Fanuc KAREL source: KT00592.KL

PROGRAM KT00592
%NOLOCKGROUP
VAR
  I1: INTEGER
  S2: STRING[80]
  OUT: STRING[80]
BEGIN
  I1 = 2
    S2 = 'B'
  OUT = I1 + S2
END KT00592
